ABB RAPID module: module1.mod

MODULE Module1
    CONST robtarget Target_10:=[[696.368666894,0,780.682032303],[0.5,0,0.866025404,0],[0,0,0,0],[9E+09,9E+09,9E+09,9E+09,9E+09,9E+09]];
    CONST robtarget Target_20:=[[527.565392707,415.534143375,54.915308258],[0.005711555,-0.000101498,0.999983683,-0.000032209],[0,-1,0,0],[9E+09,9E+09,9E+09,9E+09,9E+09,9E+09]];
    !***********************************************************
    !
    ! Module:  Module1
    !
    ! Description:
    !   Experiment to move a chess piece.
    !
    ! Author: John Cortez
    !
    ! Version: 1.0
    !
    !***********************************************************


    !***********************************************************
    !
    ! Procedure main
    !
    !   This is the entry point of your program
    !
    !***********************************************************
    PROC main()
        !Add your code here
    ENDPROC
    PROC Path_10()
        MoveL Target_10,v1000,z100,Servo\WObj:=wobj0;
        MoveL Target_20,v1000,z100,Servo\WObj:=wobj0;
    ENDPROC
ENDMODULE
